(* IEC 61131-3 sources: rusty/tests/lit/single/type_promotion/comparison, 11 files *)

(* ---- compare_guards.st ---- *)
// RUN: %COMPILE %s && %RUN | %CHECK %s
// Compares whose result does not depend on the signedness of the predicate.
FUNCTION main : DINT
    VAR
        ud : UDINT := 4000000000;
        ud2 : UDINT := 4000000000;
        ud5 : UDINT := 5;
        ul : ULINT := 18446744073709551615;
        us : USINT := 200;
        us2 : USINT := 100;
        ui : UINT := 60000;
        l1 : LINT := 1;
        sm1 : SINT := -1;
        dm10 : DINT := -10;
    END_VAR

    // Equality on values from the signed midpoint on
    printf('UDINT = UDINT = %d$N', ud = ud2);               // CHECK: UDINT = UDINT = 1
    printf('UDINT <> 5 = %d$N', ud <> ud5);                 // CHECK-NEXT: UDINT <> 5 = 1
    printf('ULINT = max = %d$N', ul = 18446744073709551615);    // CHECK-NEXT: ULINT = max = 1

    // Narrow unsigned types are widened to DINT before the compare
    printf('USINT 200 > USINT 100 = %d$N', us > us2);       // CHECK-NEXT: USINT 200 > USINT 100 = 1
    printf('UINT 60000 > 2 = %d$N', ui > 2);                // CHECK-NEXT: UINT 60000 > 2 = 1
    printf('USINT 200 > SINT -1 = %d$N', us > sm1);         // CHECK-NEXT: USINT 200 > SINT -1 = 1

    // Small unsigned values
    printf('UDINT 5 < 10 = %d$N', ud5 < 10);                // CHECK-NEXT: UDINT 5 < 10 = 1
    printf('UDINT 5 < UDINT 4e9 = %d$N', ud5 < ud);         // CHECK-NEXT: UDINT 5 < UDINT 4e9 = 1

    // A wider signed operand holds both values
    printf('UDINT 4e9 > LINT 1 = %d$N', ud > l1);           // CHECK-NEXT: UDINT 4e9 > LINT 1 = 1
    printf('UDINT 4e9 > 16#8000_0000 = %d$N', ud > 16#8000_0000);  // CHECK-NEXT: UDINT 4e9 > 16#8000_0000 = 1

    // Negative signed operands next to unsigned values
    printf('UDINT 5 > -1 = %d$N', ud5 > -1);                // CHECK-NEXT: UDINT 5 > -1 = 1
    printf('UDINT 5 > SINT -1 = %d$N', ud5 > sm1);          // CHECK-NEXT: UDINT 5 > SINT -1 = 1
    printf('DINT -10 < UDINT 5 = %d$N', dm10 < ud5);        // CHECK-NEXT: DINT -10 < UDINT 5 = 1

    // TIME, DATE and TOD below 2^31
    printf('T#1h > T#1s = %d$N', T#1h > T#1s);              // CHECK-NEXT: T#1h > T#1s = 1
    printf('TOD#23:00 > TOD#01:00 = %d$N', TOD#23:00:00 > TOD#01:00:00);  // CHECK-NEXT: TOD#23:00 > TOD#01:00 = 1
    printf('D#2020 > D#2010 = %d$N', D#2020-01-01 > D#2010-01-01);        // CHECK-NEXT: D#2020 > D#2010 = 1
    printf('LTIME#25d > LTIME#1s = %d$N', LTIME#25d > LTIME#1s);          // CHECK-NEXT: LTIME#25d > LTIME#1s = 1
END_FUNCTION

(* ---- mixed_signedness_equality.st ---- *)
// RUN: %COMPILE %s && %RUN | %CHECK %s
// XFAIL: *
// A negative signed operand and a UDINT or ULINT maximum have the same bit pattern, and = and <> compare the bits, not the values.
FUNCTION main : DINT
    VAR
        sm1 : SINT := -1;
        im1 : INT := -1;
        dm1 : DINT := -1;
        lm1 : LINT := -1;
        udmax : UDINT := 4294967295;
        ulmax : ULINT := 18446744073709551615;
    END_VAR

    printf('SINT -1 = UDINT max = %d$N', sm1 = udmax);      // CHECK: SINT -1 = UDINT max = 0
    printf('DINT -1 = UDINT max = %d$N', dm1 = udmax);      // CHECK-NEXT: DINT -1 = UDINT max = 0
    printf('DINT -1 <> UDINT max = %d$N', dm1 <> udmax);    // CHECK-NEXT: DINT -1 <> UDINT max = 1
    printf('INT -1 = ULINT max = %d$N', im1 = ulmax);       // CHECK-NEXT: INT -1 = ULINT max = 0
    printf('LINT -1 = ULINT max = %d$N', lm1 = ulmax);      // CHECK-NEXT: LINT -1 = ULINT max = 0
    printf('ULINT max <> LINT -1 = %d$N', ulmax <> lm1);    // CHECK-NEXT: ULINT max <> LINT -1 = 1
END_FUNCTION

(* ---- mixed_signedness_variables.st ---- *)
// RUN: %COMPILE %s && %RUN | %CHECK %s
// XFAIL: *
// A signed operand next to a UDINT or ULINT operand of the same or larger width makes the compare signed,
// so an unsigned value from the signed midpoint on compares as negative.
FUNCTION main : DINT
    VAR
        s5 : SINT := 5;
        d5 : DINT := 5;
        l5 : LINT := 5;
        sm1 : SINT := -1;
        dm1 : DINT := -1;
        lm1 : LINT := -1;
        i2 : INT := 2;
        d2 : DINT := 2;
        l2 : LINT := 2;
        udmax : UDINT := 4294967295;
        ulmax : ULINT := 18446744073709551615;
    END_VAR

    // Signed value below a UDINT maximum
    printf('SINT 5 < UDINT max = %d$N', s5 < udmax);        // CHECK: SINT 5 < UDINT max = 1
    printf('DINT 5 < UDINT max = %d$N', d5 < udmax);        // CHECK-NEXT: DINT 5 < UDINT max = 1
    printf('DINT -1 < UDINT max = %d$N', dm1 < udmax);      // CHECK-NEXT: DINT -1 < UDINT max = 1

    // Signed value below a ULINT maximum
    printf('DINT 5 < ULINT max = %d$N', d5 < ulmax);        // CHECK-NEXT: DINT 5 < ULINT max = 1
    printf('LINT 5 < ULINT max = %d$N', l5 < ulmax);        // CHECK-NEXT: LINT 5 < ULINT max = 1
    printf('LINT -1 < ULINT max = %d$N', lm1 < ulmax);      // CHECK-NEXT: LINT -1 < ULINT max = 1
    printf('SINT -1 < ULINT max = %d$N', sm1 < ulmax);      // CHECK-NEXT: SINT -1 < ULINT max = 1

    // Unsigned maximum on the left
    printf('UDINT max > DINT 2 = %d$N', udmax > d2);        // CHECK-NEXT: UDINT max > DINT 2 = 1
    printf('UDINT max > SINT -1 = %d$N', udmax > sm1);      // CHECK-NEXT: UDINT max > SINT -1 = 1
    printf('ULINT max > LINT 2 = %d$N', ulmax > l2);        // CHECK-NEXT: ULINT max > LINT 2 = 1
    printf('ULINT max > DINT -1 = %d$N', ulmax > dm1);      // CHECK-NEXT: ULINT max > DINT -1 = 1
    printf('ULINT max < INT 2 = %d$N', ulmax < i2);         // CHECK-NEXT: ULINT max < INT 2 = 0
END_FUNCTION

(* ---- mixed_width_unsigned_variables.st ---- *)
// RUN: %COMPILE %s && %RUN | %CHECK %s
// Two unsigned operands of different widths are promoted to the wider UDINT or ULINT and then compared unsigned.
FUNCTION main : DINT
    VAR
        us5 : USINT := 5;
        ui5 : UINT := 5;
        ud5 : UDINT := 5;
        us2 : USINT := 2;
        ui2 : UINT := 2;
        ud2 : UDINT := 2;
        udmax : UDINT := 4294967295;
        ulmax : ULINT := 18446744073709551615;
    END_VAR

    // Narrow operand next to a UDINT maximum
    printf('USINT 5 < UDINT max = %d$N', us5 < udmax);      // CHECK: USINT 5 < UDINT max = 1
    printf('UINT 5 < UDINT max = %d$N', ui5 < udmax);       // CHECK-NEXT: UINT 5 < UDINT max = 1
    printf('UDINT max > USINT 2 = %d$N', udmax > us2);      // CHECK-NEXT: UDINT max > USINT 2 = 1
    printf('UDINT max > UINT 2 = %d$N', udmax > ui2);       // CHECK-NEXT: UDINT max > UINT 2 = 1

    // Narrow operand next to a ULINT maximum
    printf('USINT 5 < ULINT max = %d$N', us5 < ulmax);      // CHECK-NEXT: USINT 5 < ULINT max = 1
    printf('ULINT max > UINT 2 = %d$N', ulmax > ui2);       // CHECK-NEXT: ULINT max > UINT 2 = 1

    // UDINT operand next to a ULINT maximum
    printf('UDINT 5 < ULINT max = %d$N', ud5 < ulmax);      // CHECK-NEXT: UDINT 5 < ULINT max = 1
    printf('ULINT max > UDINT 2 = %d$N', ulmax > ud2);      // CHECK-NEXT: ULINT max > UDINT 2 = 1
END_FUNCTION

(* ---- time_and_date_after_midpoint.st ---- *)
// RUN: %COMPILE %s && %RUN | %CHECK %s
// TIME, DATE and DT are unsigned 32-bit values and compare unsigned, so values from 2^31 on compare as large.
FUNCTION main : DINT
    VAR
        long_time : TIME := T#25d;
        short_time : TIME := T#1h;
        later : DT := DT#2038-01-19-03:14:08;
        earlier : DT := DT#2038-01-19-03:14:07;
        future : DATE := D#2040-01-01;
        past : DATE := D#2020-01-01;
    END_VAR

    // TIME above about 24.8 days
    printf('T#25d > T#1h = %d$N', long_time > short_time);  // CHECK: T#25d > T#1h = 1
    printf('T#1h < T#25d = %d$N', short_time < long_time);  // CHECK-NEXT: T#1h < T#25d = 1
    printf('T#24d21h > T#24d20h = %d$N', T#24d21h > T#24d20h);  // CHECK-NEXT: T#24d21h > T#24d20h = 1

    // DT and DATE after 2038-01-19 03:14:07
    printf('later > earlier = %d$N', later > earlier);      // CHECK-NEXT: later > earlier = 1
    printf('2040 > 2020 = %d$N', future > past);            // CHECK-NEXT: 2040 > 2020 = 1
    printf('2020 >= 2040 = %d$N', past >= future);          // CHECK-NEXT: 2020 >= 2040 = 0
END_FUNCTION

(* ---- udint_variables.st ---- *)
// RUN: %COMPILE %s && %RUN | %CHECK %s
// A relational compare of two UDINT values is unsigned, so a value from the signed midpoint on compares as large.
FUNCTION main : DINT
    VAR
        hi : UDINT := 4000000000;
        lo : UDINT := 5;
        mid : UDINT := 2147483648;
        below : UDINT := 2147483647;
        result : BOOL;
    END_VAR

    // Every relational operator, both operand orders
    printf('hi > lo = %d$N', hi > lo);             // CHECK: hi > lo = 1
    printf('hi >= lo = %d$N', hi >= lo);           // CHECK-NEXT: hi >= lo = 1
    printf('hi < lo = %d$N', hi < lo);             // CHECK-NEXT: hi < lo = 0
    printf('hi <= lo = %d$N', hi <= lo);           // CHECK-NEXT: hi <= lo = 0
    printf('lo < hi = %d$N', lo < hi);             // CHECK-NEXT: lo < hi = 1
    printf('lo <= hi = %d$N', lo <= hi);           // CHECK-NEXT: lo <= hi = 1
    printf('lo > hi = %d$N', lo > hi);             // CHECK-NEXT: lo > hi = 0
    printf('lo >= hi = %d$N', lo >= hi);           // CHECK-NEXT: lo >= hi = 0

    // The two values next to the signed midpoint
    printf('mid > below = %d$N', mid > below);     // CHECK-NEXT: mid > below = 1

    // A typed literal operand of the same type
    printf('hi > UDINT#5 = %d$N', hi > UDINT#5);  // CHECK-NEXT: hi > UDINT#5 = 1

    // The compare as a stored value and as a condition
    result := hi > lo;
    printf('stored = %d$N', result);               // CHECK-NEXT: stored = 1
    IF hi > lo THEN
        printf('IF taken$N');                      // CHECK-NEXT: IF taken
    ELSE
        printf('IF not taken$N');
    END_IF
END_FUNCTION

(* ---- ulint_variables.st ---- *)
// RUN: %COMPILE %s && %RUN | %CHECK %s
// A relational compare of two ULINT values is unsigned, so a value from the signed midpoint on compares as large.
FUNCTION main : DINT
    VAR
        hi : ULINT := 18446744073709551615;
        lo : ULINT := 5;
        mid : ULINT := 9223372036854775808;
        below : ULINT := 9223372036854775807;
        result : BOOL;
    END_VAR

    // Every relational operator, both operand orders
    printf('hi > lo = %d$N', hi > lo);             // CHECK: hi > lo = 1
    printf('hi >= lo = %d$N', hi >= lo);           // CHECK-NEXT: hi >= lo = 1
    printf('hi < lo = %d$N', hi < lo);             // CHECK-NEXT: hi < lo = 0
    printf('hi <= lo = %d$N', hi <= lo);           // CHECK-NEXT: hi <= lo = 0
    printf('lo < hi = %d$N', lo < hi);             // CHECK-NEXT: lo < hi = 1
    printf('lo <= hi = %d$N', lo <= hi);           // CHECK-NEXT: lo <= hi = 1
    printf('lo > hi = %d$N', lo > hi);             // CHECK-NEXT: lo > hi = 0
    printf('lo >= hi = %d$N', lo >= hi);           // CHECK-NEXT: lo >= hi = 0

    // The two values next to the signed midpoint
    printf('mid > below = %d$N', mid > below);     // CHECK-NEXT: mid > below = 1

    // A typed literal operand of the same type
    printf('hi > ULINT#5 = %d$N', hi > ULINT#5);  // CHECK-NEXT: hi > ULINT#5 = 1

    // The compare as a stored value and as a condition
    result := hi > lo;
    printf('stored = %d$N', result);               // CHECK-NEXT: stored = 1
    IF hi > lo THEN
        printf('IF taken$N');                      // CHECK-NEXT: IF taken
    ELSE
        printf('IF not taken$N');
    END_IF
END_FUNCTION

(* ---- unsigned_comparison_functions.st ---- *)
// RUN: %COMPILE %s && %RUN | %CHECK %s
// The comparison functions compare two UDINT values unsigned, as the operators do.
FUNCTION main : DINT
    VAR
        hi : UDINT := 4000000000;
        mid : UDINT := 3000000000;
        lo : UDINT := 5;
    END_VAR

    printf('GT(hi, lo) = %d$N', GT(hi, lo));                // CHECK: GT(hi, lo) = 1
    printf('GE(hi, lo) = %d$N', GE(hi, lo));                // CHECK-NEXT: GE(hi, lo) = 1
    printf('LT(lo, hi) = %d$N', LT(lo, hi));                // CHECK-NEXT: LT(lo, hi) = 1
    printf('LE(lo, hi) = %d$N', LE(lo, hi));                // CHECK-NEXT: LE(lo, hi) = 1
    printf('GT(hi, mid, lo) = %d$N', GT(hi, mid, lo));      // CHECK-NEXT: GT(hi, mid, lo) = 1
    printf('LT(lo, mid, hi) = %d$N', LT(lo, mid, hi));      // CHECK-NEXT: LT(lo, mid, hi) = 1
    printf('MAX(hi, lo) = %u$N', MAX(hi, lo));              // CHECK-NEXT: MAX(hi, lo) = 4000000000
    printf('MIN(hi, lo) = %u$N', MIN(hi, lo));              // CHECK-NEXT: MIN(hi, lo) = 5
    printf('LIMIT(lo, hi, mid) = %u$N', LIMIT(lo, hi, mid));    // CHECK-NEXT: LIMIT(lo, hi, mid) = 3000000000
END_FUNCTION

(* ---- unsigned_with_negative_literal.st ---- *)
// RUN: %COMPILE %s && %RUN | %CHECK %s
// XFAIL: *
// A negative literal next to a UDINT or ULINT maximum compares signed, so the maximum reads as -1.
FUNCTION main : DINT
    VAR
        udmax : UDINT := 4294967295;
        ulmax : ULINT := 18446744073709551615;
    END_VAR

    // Relational compares
    printf('UDINT max > -1 = %d$N', udmax > -1);            // CHECK: UDINT max > -1 = 1
    printf('ULINT max > -1 = %d$N', ulmax > -1);            // CHECK-NEXT: ULINT max > -1 = 1
    printf('-1 < UDINT max = %d$N', -1 < udmax);            // CHECK-NEXT: -1 < UDINT max = 1
    printf('-1 < ULINT max = %d$N', -1 < ulmax);            // CHECK-NEXT: -1 < ULINT max = 1

    // Equality
    printf('UDINT max = -1 = %d$N', udmax = -1);            // CHECK-NEXT: UDINT max = -1 = 0
    printf('ULINT max = -1 = %d$N', ulmax = -1);            // CHECK-NEXT: ULINT max = -1 = 0
    printf('UDINT max <> -1 = %d$N', udmax <> -1);          // CHECK-NEXT: UDINT max <> -1 = 1
END_FUNCTION

(* ---- unsigned_with_untyped_literal.st ---- *)
// RUN: %COMPILE %s && %RUN | %CHECK %s
// An untyped integer literal takes the type of a UDINT or ULINT operand, so the compare is unsigned.
FUNCTION main : DINT
    VAR
        ud : UDINT := 4000000000;
        ul : ULINT := 18446744073709551615;
    END_VAR

    // Literal on the right
    printf('UDINT > 5 = %d$N', ud > 5);                     // CHECK: UDINT > 5 = 1
    printf('UDINT >= 2147483647 = %d$N', ud >= 2147483647); // CHECK-NEXT: UDINT >= 2147483647 = 1
    printf('UDINT < 5 = %d$N', ud < 5);                     // CHECK-NEXT: UDINT < 5 = 0
    printf('UDINT < 0 = %d$N', ud < 0);                     // CHECK-NEXT: UDINT < 0 = 0
    printf('ULINT > 1 = %d$N', ul > 1);                     // CHECK-NEXT: ULINT > 1 = 1
    printf('ULINT > 3000000000 = %d$N', ul > 3000000000);   // CHECK-NEXT: ULINT > 3000000000 = 1

    // Literal on the left
    printf('5 < UDINT = %d$N', 5 < ud);                     // CHECK-NEXT: 5 < UDINT = 1
    printf('1 < ULINT = %d$N', 1 < ul);                     // CHECK-NEXT: 1 < ULINT = 1
END_FUNCTION

(* ---- literal_by_declaration_section.st ---- *)
// RUN: %COMPILE %s && %RUN | %CHECK %s
// A compare of a UDINT or ULINT operand with an untyped literal is unsigned, wherever the operand is declared.
VAR_GLOBAL
    g : UDINT := 4294967295;
END_VAR

VAR_GLOBAL CONSTANT
    gc : ULINT := 18446744073709551615;
END_VAR

FUNCTION_BLOCK probe
    VAR_INPUT
        i : UDINT;
    END_VAR
    VAR_INPUT CONSTANT
        ic : UDINT := 4294967295;
    END_VAR
    VAR_IN_OUT
        io : ULINT;
    END_VAR
    VAR_OUTPUT
        o : UDINT;
    END_VAR
    VAR
        m : ULINT := 18446744073709551615;
    END_VAR
    VAR CONSTANT
        c : UDINT := 4294967295;
    END_VAR
    VAR_TEMP
        t : UDINT;
    END_VAR

    o := 4294967295;
    t := 4294967295;
    printf('VAR_INPUT > 16#7FFFFFFF = %d$N', i > 16#7FFFFFFF);
    printf('VAR_INPUT CONSTANT < 0 = %d$N', ic < 0);
    printf('VAR_IN_OUT > 16#7FFFFFFF = %d$N', io > 16#7FFFFFFF);
    printf('VAR_OUTPUT < 0 = %d$N', o < 0);
    printf('VAR > 3000000000 = %d$N', m > 3000000000);
    printf('VAR CONSTANT > 16#7FFFFFFF = %d$N', c > 16#7FFFFFFF);
    printf('VAR_TEMP < 0 = %d$N', t < 0);
    printf('VAR_GLOBAL > 16#7FFFFFFF = %d$N', g > 16#7FFFFFFF);
    printf('VAR_GLOBAL CONSTANT < 0 = %d$N', gc < 0);
END_FUNCTION_BLOCK

FUNCTION main : DINT
    VAR
        inst : probe;
        v : ULINT := 18446744073709551615;
    END_VAR

    inst(i := 4294967295, io := v);
    // CHECK: VAR_INPUT > 16#7FFFFFFF = 1
    // CHECK-NEXT: VAR_INPUT CONSTANT < 0 = 0
    // CHECK-NEXT: VAR_IN_OUT > 16#7FFFFFFF = 1
    // CHECK-NEXT: VAR_OUTPUT < 0 = 0
    // CHECK-NEXT: VAR > 3000000000 = 1
    // CHECK-NEXT: VAR CONSTANT > 16#7FFFFFFF = 1
    // CHECK-NEXT: VAR_TEMP < 0 = 0
    // CHECK-NEXT: VAR_GLOBAL > 16#7FFFFFFF = 1
    // CHECK-NEXT: VAR_GLOBAL CONSTANT < 0 = 0
END_FUNCTION
